(* Logix 5000 project; controller _1407974_PSG_7315 vendor 1 type 14 code 154 rev 20.11; software revision 20.06; part 2 of 4 *)
(* tags used below, declared in another part *)
   AI_L_2_1_FW_Pressure : Analog_Input;
   AI_R_2_0_Pure_Steam_Temperature : Analog_Input;
   Alarm_Emergency_Stop : ALIAS FOR Alarms_Warnings.Latch_Bit[0].0;
   Alarm_Emergency_Stop_Ack : ALIAS FOR Alarms_Warnings.Ack[0].0;
   Alarm_Pure_Steam_High_Temp_Timer : TIMER;
   Alarm_Pure_Steam_High_Temperature : ALIAS FOR Alarms_Warnings.Latch_Bit[0].4;
   Alarm_Pure_Steam_High_Temperature_Ack : ALIAS FOR Alarms_Warnings.Ack[0].4;
   Alarm_Pure_Steam_Temp_Error_Timer : TIMER;
   Alarm_Rupture_Disk_Failure : ALIAS FOR Alarms_Warnings.Latch_Bit[0].1;
   Alarm_Rupture_Disk_Failure_Timer : TIMER;
   Alarm_Rupture_Disk_Faiure_Ack : ALIAS FOR Alarms_Warnings.Ack[0].1;
   Alarm_Separator_High_Level : ALIAS FOR Alarms_Warnings.Latch_Bit[0].2;
   Alarm_Separator_High_Level_Ack : ALIAS FOR Alarms_Warnings.Ack[0].2;
   Alarm_Separator_High_Level_Timer : TIMER;
   Alarm_Separator_Low_Level : ALIAS FOR Alarms_Warnings.Latch_Bit[0].3;
   Alarm_Separator_Low_Level_Ack : ALIAS FOR Alarms_Warnings.Ack[0].3;
   Alarm_Separator_Low_Level_Timer_A : TIMER;
   Alarm_Separator_Low_Level_Timer_B : TIMER;
   Alarms_Warnings : AW;
   AO_L_3_0_VFD_SPEED : Analog_Output;
   AO_R_4_0_Pure_Steam_Temperature : Analog_Output;
   Calculated_CV_Max_Value : REAL;
   Condensed_Pure_Steam_Warrnings_Disabled : Latched_Push_Button;
   Cooling_State_Latch_Timer : TIMER;
   Cooling_Status_Debounce_Timer : TIMER;
   DI_L_1_0_Emergency_Stop_Relay : ALIAS FOR DI_Local_1.0;
   DI_R_1_0_Hi_Hi_Level_LSHH_1950 : ALIAS FOR DI_Remote_1.0;
   DI_R_1_1_Hi_Level_LSH_1950 : ALIAS FOR DI_Remote_1.1;
   DI_R_1_2_Mid_Level_LSM_1950 : ALIAS FOR DI_Remote_1.2;
   DI_R_1_3_Low_Level_LSL_1950 : ALIAS FOR DI_Remote_1.3;
   DI_R_1_5_Burst_Disk_Sensor_PSH_5820 : ALIAS FOR DI_Remote_1.5;
   DO_L_1_0_Alarm_Relay_Coil : Discrete_Out;
   DO_L_1_10_Available : Discrete_Out;
   DO_L_1_11_Available : Discrete_Out;
   DO_L_1_12_Available : Discrete_Out;
   DO_L_1_13_Available : Discrete_Out;
   DO_L_1_14_Feed_Water_Pump_Contactor : Discrete_Out;
   DO_L_1_15_Feed_Water_Pump_On_Light : Discrete_Out;
   DO_L_1_1_Alarm_Horn : Discrete_Out;
   DO_L_1_2_Alarm_Light : Discrete_Out;
   DO_L_1_3_Ready_Light : Discrete_Out;
   DO_L_1_4_Running_Light : Discrete_Out;
   DO_L_1_5_Hour_Meter : Discrete_Out;
   DO_L_1_6_Available : Discrete_Out;
   DO_L_1_7_Available : Discrete_Out;
   DO_L_1_8_Available : Discrete_Out;
   DO_L_1_9_Available : Discrete_Out;
   DO_R_3_0_Pure_Steam_Temp_Control_YV_4110 : Discrete_Out;
   DO_R_3_1_Primary_Level_Control_YV_4760 : Discrete_Out;
   DO_R_3_2_Secondary_Level_Control_YV_4770 : Discrete_Out;
   DO_R_3_3_Coolant_Shutoff_FCV_3025 : Discrete_Out;
   DO_R_3_4_Degasser_Vent_YV_4255 : Discrete_Out;
   DO_R_3_5_FDW_TR : Discrete_Out;
   DO_R_3_6_Available : Discrete_Out;
   DO_R_3_7_Available : Discrete_Out;
   Feedwater_Pressure_PID : PID;
   Feedwater_Pressure_PID_Auto_Mode : Push_Button;
   Feedwater_Pressure_PID_Manual_Mode : Push_Button;
   Lamp_Test : Push_Button;
   Local_Remote : Latched_Push_Button;
   Low_Level_Latch : BOOL;
   Maintenance_Mode : Latched_Push_Button;
   Network_Start : BOOL;
   Network_Stop : BOOL;
   OIT : OIT_Connections;
   PID_Auto_Mode : Push_Button;
   PID_CV_Max_Value_Initialize : BOOL;
   PID_Loop_Trigger_Timer : TIMER;
   PID_Manual_Mode : Push_Button;
   PID_Ramp_Timer : TIMER;
   PS_Temp_GEQ_SetPoint_Minus_5_Deg : BOOL;
   PS_Temp_Setpoint_Minus_5_Deg : REAL;
   Pure_Steam_Temp_Output_Clamp : BOOL;
   Pure_Steam_Temperature : PID;
   Start : Push_Button;
   Stop : Push_Button;
   Unit_Hot : BOOL;
   Unit_Status : Unit_Status;
(* MainProgram, continued *)

ROUTINE _050_Maintenance   (* ladder *)
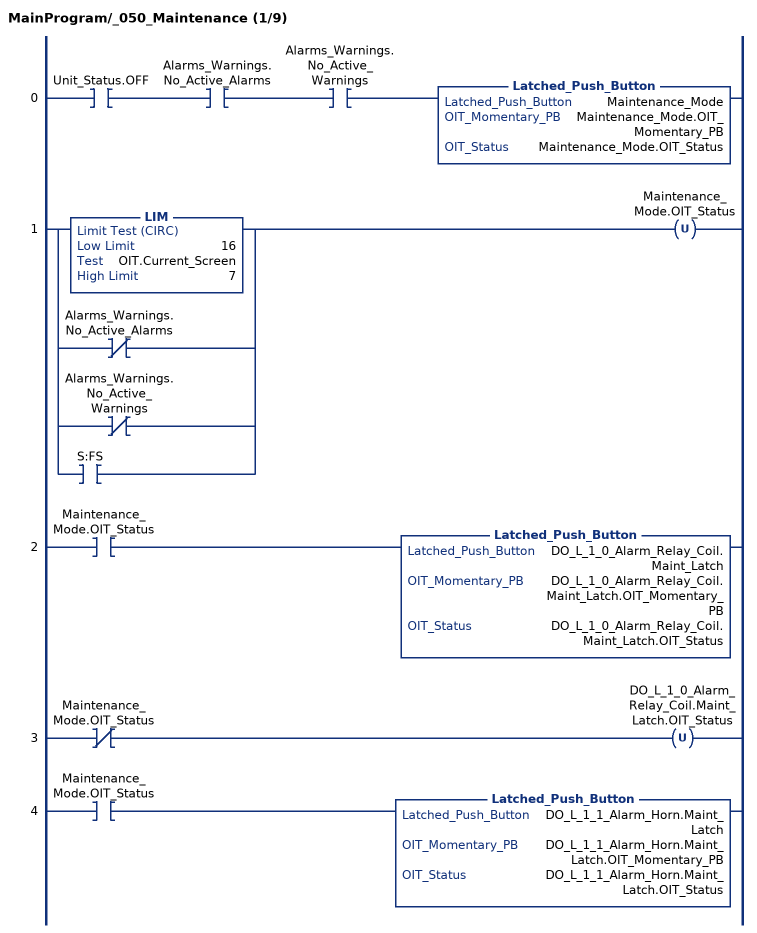
   0: XIC(Unit_Status.OFF)XIC(Alarms_Warnings.No_Active_Alarms)XIC(Alarms_Warnings.No_Active_Warnings)Latched_Push_Button(Maintenance_Mode,Maintenance_Mode.OIT_Momentary_PB,Maintenance_Mode.OIT_Status);
   1: [LIM(16,OIT.Current_Screen,7) ,XIO(Alarms_Warnings.No_Active_Alarms) ,XIO(Alarms_Warnings.No_Active_Warnings) ,XIC(S:FS) ]OTU(Maintenance_Mode.OIT_Status);
   2: XIC(Maintenance_Mode.OIT_Status)Latched_Push_Button(DO_L_1_0_Alarm_Relay_Coil.Maint_Latch,DO_L_1_0_Alarm_Relay_Coil.Maint_Latch.OIT_Momentary_PB,DO_L_1_0_Alarm_Relay_Coil.Maint_Latch.OIT_Status);
   3: XIO(Maintenance_Mode.OIT_Status)OTU(DO_L_1_0_Alarm_Relay_Coil.Maint_Latch.OIT_Status);
   4: XIC(Maintenance_Mode.OIT_Status)Latched_Push_Button(DO_L_1_1_Alarm_Horn.Maint_Latch,DO_L_1_1_Alarm_Horn.Maint_Latch.OIT_Momentary_PB,DO_L_1_1_Alarm_Horn.Maint_Latch.OIT_Status);
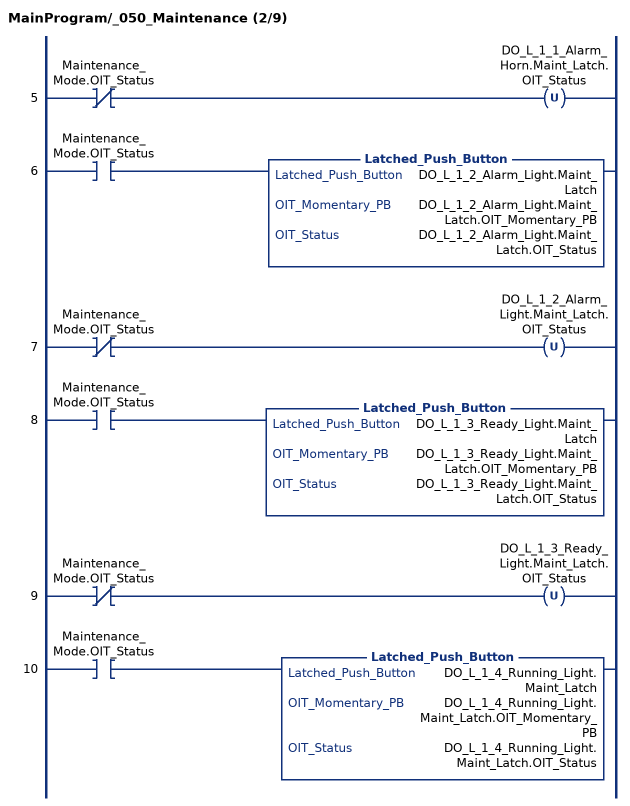
   5: XIO(Maintenance_Mode.OIT_Status)OTU(DO_L_1_1_Alarm_Horn.Maint_Latch.OIT_Status);
   6: XIC(Maintenance_Mode.OIT_Status)Latched_Push_Button(DO_L_1_2_Alarm_Light.Maint_Latch,DO_L_1_2_Alarm_Light.Maint_Latch.OIT_Momentary_PB,DO_L_1_2_Alarm_Light.Maint_Latch.OIT_Status);
   7: XIO(Maintenance_Mode.OIT_Status)OTU(DO_L_1_2_Alarm_Light.Maint_Latch.OIT_Status);
   8: XIC(Maintenance_Mode.OIT_Status)Latched_Push_Button(DO_L_1_3_Ready_Light.Maint_Latch,DO_L_1_3_Ready_Light.Maint_Latch.OIT_Momentary_PB,DO_L_1_3_Ready_Light.Maint_Latch.OIT_Status);
   9: XIO(Maintenance_Mode.OIT_Status)OTU(DO_L_1_3_Ready_Light.Maint_Latch.OIT_Status);
   10: XIC(Maintenance_Mode.OIT_Status)Latched_Push_Button(DO_L_1_4_Running_Light.Maint_Latch,DO_L_1_4_Running_Light.Maint_Latch.OIT_Momentary_PB,DO_L_1_4_Running_Light.Maint_Latch.OIT_Status);
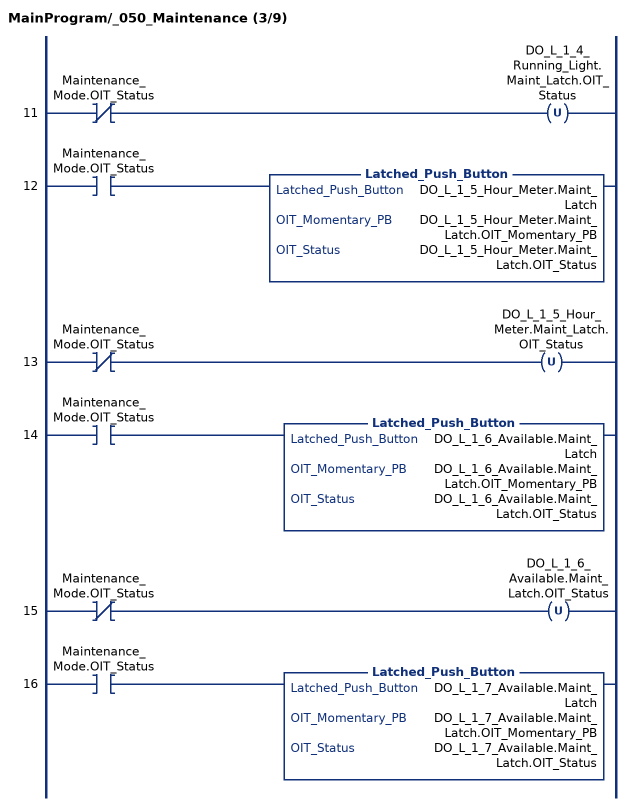
   11: XIO(Maintenance_Mode.OIT_Status)OTU(DO_L_1_4_Running_Light.Maint_Latch.OIT_Status);
   12: XIC(Maintenance_Mode.OIT_Status)Latched_Push_Button(DO_L_1_5_Hour_Meter.Maint_Latch,DO_L_1_5_Hour_Meter.Maint_Latch.OIT_Momentary_PB,DO_L_1_5_Hour_Meter.Maint_Latch.OIT_Status);
   13: XIO(Maintenance_Mode.OIT_Status)OTU(DO_L_1_5_Hour_Meter.Maint_Latch.OIT_Status);
   14: XIC(Maintenance_Mode.OIT_Status)Latched_Push_Button(DO_L_1_6_Available.Maint_Latch,DO_L_1_6_Available.Maint_Latch.OIT_Momentary_PB,DO_L_1_6_Available.Maint_Latch.OIT_Status);
   15: XIO(Maintenance_Mode.OIT_Status)OTU(DO_L_1_6_Available.Maint_Latch.OIT_Status);
   16: XIC(Maintenance_Mode.OIT_Status)Latched_Push_Button(DO_L_1_7_Available.Maint_Latch,DO_L_1_7_Available.Maint_Latch.OIT_Momentary_PB,DO_L_1_7_Available.Maint_Latch.OIT_Status);
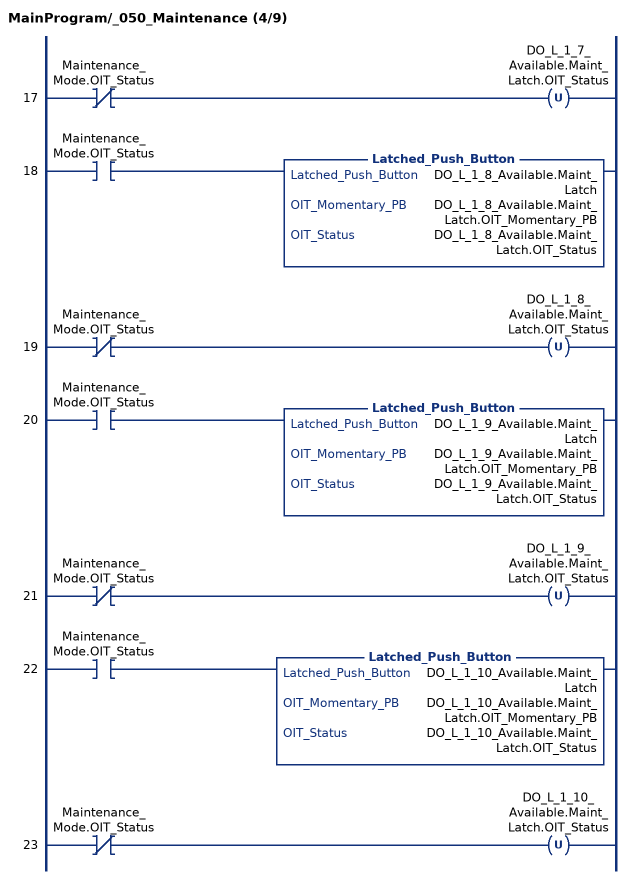
   17: XIO(Maintenance_Mode.OIT_Status)OTU(DO_L_1_7_Available.Maint_Latch.OIT_Status);
   18: XIC(Maintenance_Mode.OIT_Status)Latched_Push_Button(DO_L_1_8_Available.Maint_Latch,DO_L_1_8_Available.Maint_Latch.OIT_Momentary_PB,DO_L_1_8_Available.Maint_Latch.OIT_Status);
   19: XIO(Maintenance_Mode.OIT_Status)OTU(DO_L_1_8_Available.Maint_Latch.OIT_Status);
   20: XIC(Maintenance_Mode.OIT_Status)Latched_Push_Button(DO_L_1_9_Available.Maint_Latch,DO_L_1_9_Available.Maint_Latch.OIT_Momentary_PB,DO_L_1_9_Available.Maint_Latch.OIT_Status);
   21: XIO(Maintenance_Mode.OIT_Status)OTU(DO_L_1_9_Available.Maint_Latch.OIT_Status);
   22: XIC(Maintenance_Mode.OIT_Status)Latched_Push_Button(DO_L_1_10_Available.Maint_Latch,DO_L_1_10_Available.Maint_Latch.OIT_Momentary_PB,DO_L_1_10_Available.Maint_Latch.OIT_Status);
   23: XIO(Maintenance_Mode.OIT_Status)OTU(DO_L_1_10_Available.Maint_Latch.OIT_Status);
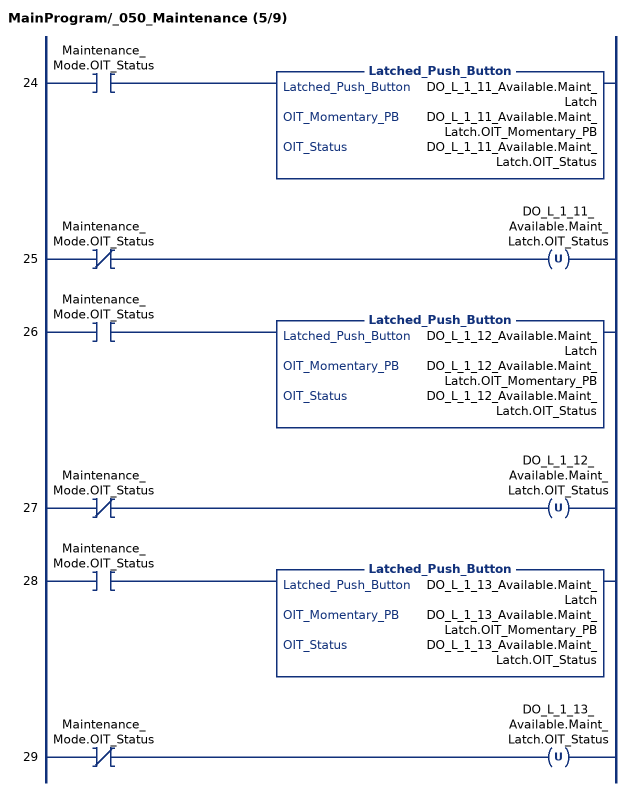
   24: XIC(Maintenance_Mode.OIT_Status)Latched_Push_Button(DO_L_1_11_Available.Maint_Latch,DO_L_1_11_Available.Maint_Latch.OIT_Momentary_PB,DO_L_1_11_Available.Maint_Latch.OIT_Status);
   25: XIO(Maintenance_Mode.OIT_Status)OTU(DO_L_1_11_Available.Maint_Latch.OIT_Status);
   26: XIC(Maintenance_Mode.OIT_Status)Latched_Push_Button(DO_L_1_12_Available.Maint_Latch,DO_L_1_12_Available.Maint_Latch.OIT_Momentary_PB,DO_L_1_12_Available.Maint_Latch.OIT_Status);
   27: XIO(Maintenance_Mode.OIT_Status)OTU(DO_L_1_12_Available.Maint_Latch.OIT_Status);
   28: XIC(Maintenance_Mode.OIT_Status)Latched_Push_Button(DO_L_1_13_Available.Maint_Latch,DO_L_1_13_Available.Maint_Latch.OIT_Momentary_PB,DO_L_1_13_Available.Maint_Latch.OIT_Status);
   29: XIO(Maintenance_Mode.OIT_Status)OTU(DO_L_1_13_Available.Maint_Latch.OIT_Status);
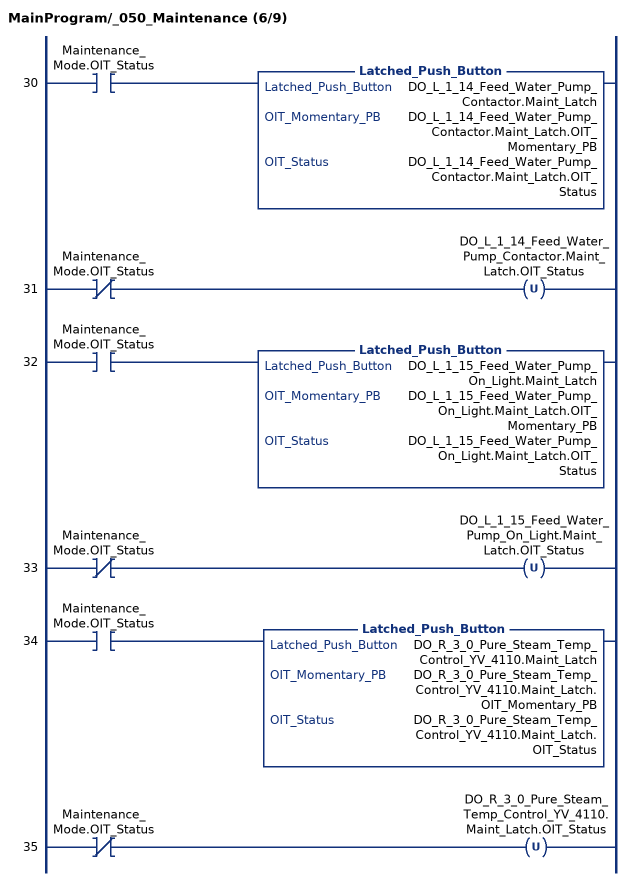
   30: XIC(Maintenance_Mode.OIT_Status)Latched_Push_Button(DO_L_1_14_Feed_Water_Pump_Contactor.Maint_Latch,DO_L_1_14_Feed_Water_Pump_Contactor.Maint_Latch.OIT_Momentary_PB,DO_L_1_14_Feed_Water_Pump_Contactor.Maint_Latch.OIT_Status);
   31: XIO(Maintenance_Mode.OIT_Status)OTU(DO_L_1_14_Feed_Water_Pump_Contactor.Maint_Latch.OIT_Status);
   32: XIC(Maintenance_Mode.OIT_Status)Latched_Push_Button(DO_L_1_15_Feed_Water_Pump_On_Light.Maint_Latch,DO_L_1_15_Feed_Water_Pump_On_Light.Maint_Latch.OIT_Momentary_PB,DO_L_1_15_Feed_Water_Pump_On_Light.Maint_Latch.OIT_Status);
   33: XIO(Maintenance_Mode.OIT_Status)OTU(DO_L_1_15_Feed_Water_Pump_On_Light.Maint_Latch.OIT_Status);
   34: XIC(Maintenance_Mode.OIT_Status)Latched_Push_Button(DO_R_3_0_Pure_Steam_Temp_Control_YV_4110.Maint_Latch,DO_R_3_0_Pure_Steam_Temp_Control_YV_4110.Maint_Latch.OIT_Momentary_PB,DO_R_3_0_Pure_Steam_Temp_Control_YV_4110.Maint_Latch.OIT_Status);
   35: XIO(Maintenance_Mode.OIT_Status)OTU(DO_R_3_0_Pure_Steam_Temp_Control_YV_4110.Maint_Latch.OIT_Status);
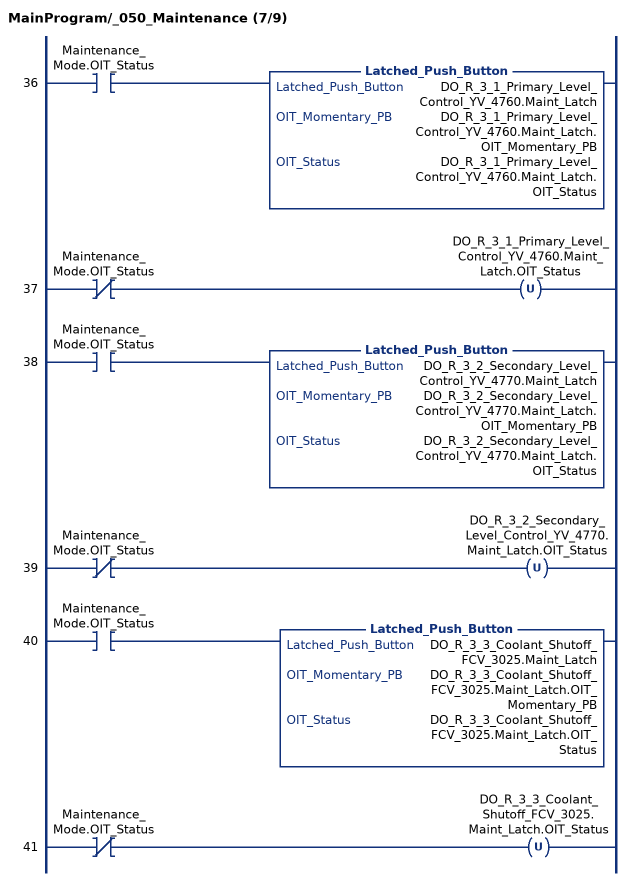
   36: XIC(Maintenance_Mode.OIT_Status)Latched_Push_Button(DO_R_3_1_Primary_Level_Control_YV_4760.Maint_Latch,DO_R_3_1_Primary_Level_Control_YV_4760.Maint_Latch.OIT_Momentary_PB,DO_R_3_1_Primary_Level_Control_YV_4760.Maint_Latch.OIT_Status);
   37: XIO(Maintenance_Mode.OIT_Status)OTU(DO_R_3_1_Primary_Level_Control_YV_4760.Maint_Latch.OIT_Status);
   38: XIC(Maintenance_Mode.OIT_Status)Latched_Push_Button(DO_R_3_2_Secondary_Level_Control_YV_4770.Maint_Latch,DO_R_3_2_Secondary_Level_Control_YV_4770.Maint_Latch.OIT_Momentary_PB,DO_R_3_2_Secondary_Level_Control_YV_4770.Maint_Latch.OIT_Status);
   39: XIO(Maintenance_Mode.OIT_Status)OTU(DO_R_3_2_Secondary_Level_Control_YV_4770.Maint_Latch.OIT_Status);
   40: XIC(Maintenance_Mode.OIT_Status)Latched_Push_Button(DO_R_3_3_Coolant_Shutoff_FCV_3025.Maint_Latch,DO_R_3_3_Coolant_Shutoff_FCV_3025.Maint_Latch.OIT_Momentary_PB,DO_R_3_3_Coolant_Shutoff_FCV_3025.Maint_Latch.OIT_Status);
   41: XIO(Maintenance_Mode.OIT_Status)OTU(DO_R_3_3_Coolant_Shutoff_FCV_3025.Maint_Latch.OIT_Status);
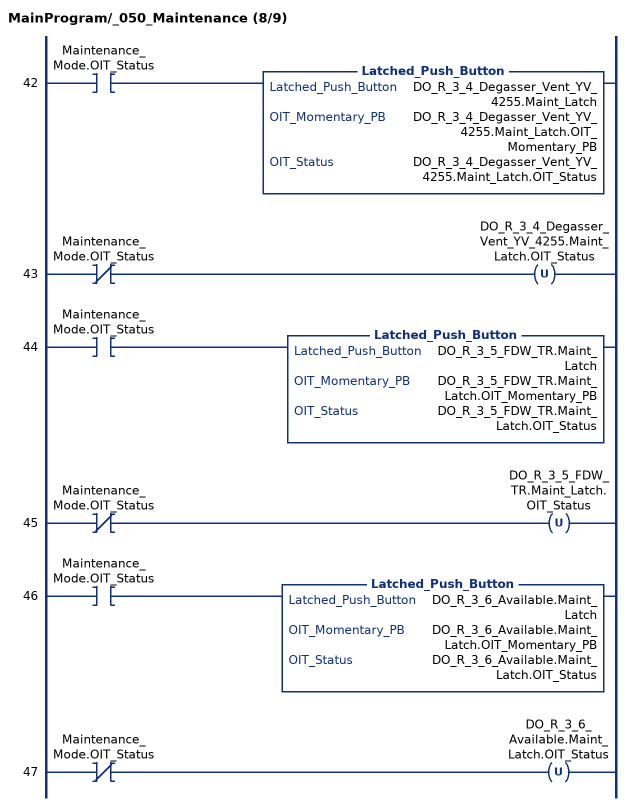
   42: XIC(Maintenance_Mode.OIT_Status)Latched_Push_Button(DO_R_3_4_Degasser_Vent_YV_4255.Maint_Latch,DO_R_3_4_Degasser_Vent_YV_4255.Maint_Latch.OIT_Momentary_PB,DO_R_3_4_Degasser_Vent_YV_4255.Maint_Latch.OIT_Status);
   43: XIO(Maintenance_Mode.OIT_Status)OTU(DO_R_3_4_Degasser_Vent_YV_4255.Maint_Latch.OIT_Status);
   44: XIC(Maintenance_Mode.OIT_Status)Latched_Push_Button(DO_R_3_5_FDW_TR.Maint_Latch,DO_R_3_5_FDW_TR.Maint_Latch.OIT_Momentary_PB,DO_R_3_5_FDW_TR.Maint_Latch.OIT_Status);
   45: XIO(Maintenance_Mode.OIT_Status)OTU(DO_R_3_5_FDW_TR.Maint_Latch.OIT_Status);
   46: XIC(Maintenance_Mode.OIT_Status)Latched_Push_Button(DO_R_3_6_Available.Maint_Latch,DO_R_3_6_Available.Maint_Latch.OIT_Momentary_PB,DO_R_3_6_Available.Maint_Latch.OIT_Status);
   47: XIO(Maintenance_Mode.OIT_Status)OTU(DO_R_3_6_Available.Maint_Latch.OIT_Status);
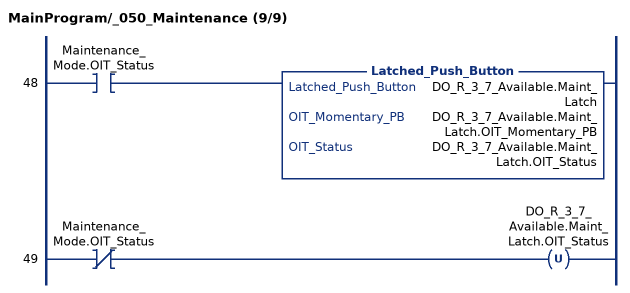
   48: XIC(Maintenance_Mode.OIT_Status)Latched_Push_Button(DO_R_3_7_Available.Maint_Latch,DO_R_3_7_Available.Maint_Latch.OIT_Momentary_PB,DO_R_3_7_Available.Maint_Latch.OIT_Status);
   49: XIO(Maintenance_Mode.OIT_Status)OTU(DO_R_3_7_Available.Maint_Latch.OIT_Status);
END_ROUTINE

ROUTINE _060_Main_Routine   (* ladder *)
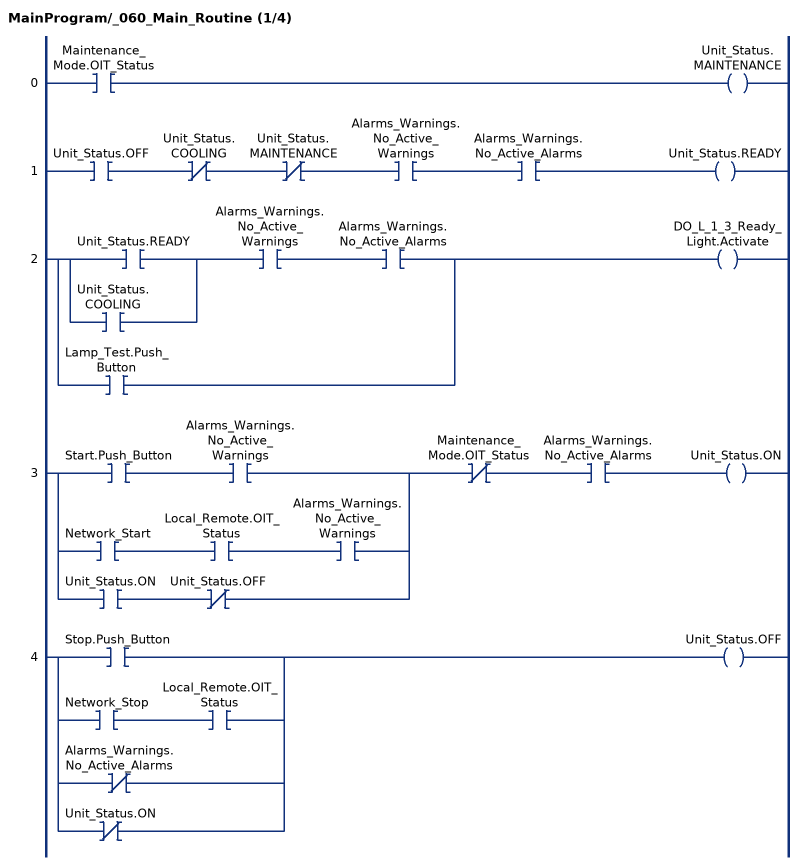
   0: XIC(Maintenance_Mode.OIT_Status)OTE(Unit_Status.MAINTENANCE);
   1: XIC(Unit_Status.OFF)XIO(Unit_Status.COOLING)XIO(Unit_Status.MAINTENANCE)XIC(Alarms_Warnings.No_Active_Warnings)XIC(Alarms_Warnings.No_Active_Alarms)OTE(Unit_Status.READY);
   2: [[XIC(Unit_Status.READY) ,XIC(Unit_Status.COOLING) ] XIC(Alarms_Warnings.No_Active_Warnings) XIC(Alarms_Warnings.No_Active_Alarms) ,XIC(Lamp_Test.Push_Button) ]OTE(DO_L_1_3_Ready_Light.Activate);
   3: [XIC(Start.Push_Button) XIC(Alarms_Warnings.No_Active_Warnings) ,XIC(Network_Start) XIC(Local_Remote.OIT_Status) XIC(Alarms_Warnings.No_Active_Warnings) ,XIC(Unit_Status.ON) XIO(Unit_Status.OFF) ]XIO(Maintenance_Mode.OIT_Status)XIC(Alarms_Warnings.No_Active_Alarms)OTE(Unit_Status.ON);
   4: [XIC(Stop.Push_Button) ,XIC(Network_Stop) XIC(Local_Remote.OIT_Status) ,XIO(Alarms_Warnings.No_Active_Alarms) ,XIO(Unit_Status.ON) ]OTE(Unit_Status.OFF);
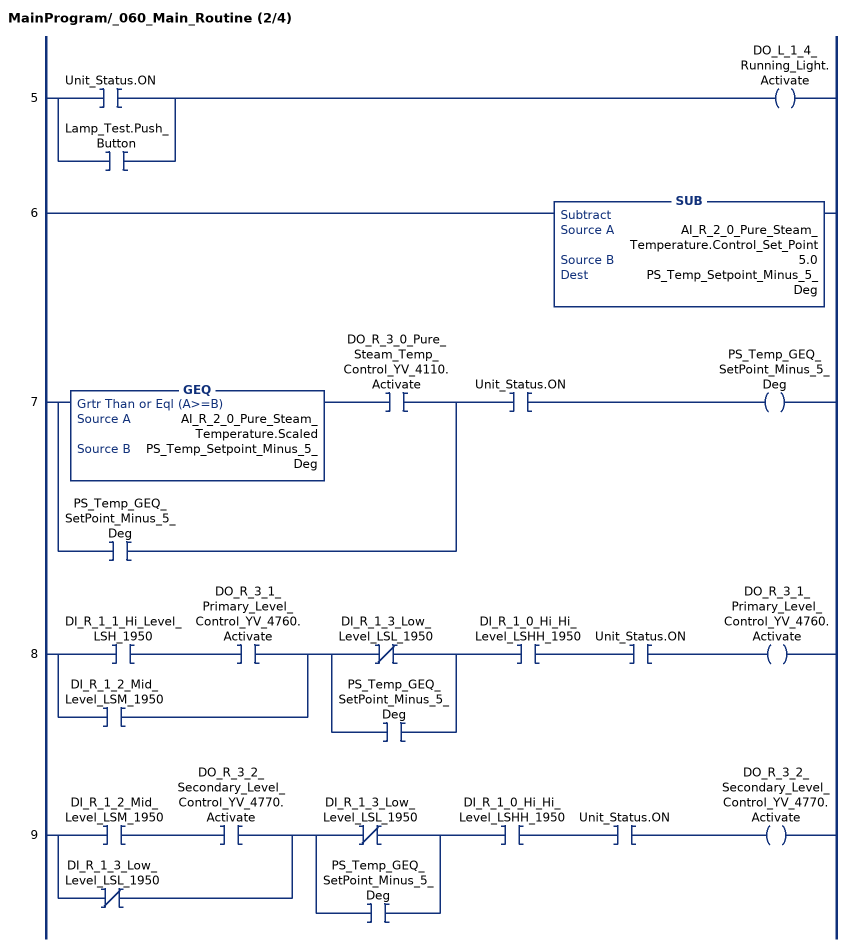
   5: [XIC(Unit_Status.ON) ,XIC(Lamp_Test.Push_Button) ]OTE(DO_L_1_4_Running_Light.Activate);
   6: SUB(AI_R_2_0_Pure_Steam_Temperature.Control_Set_Point,5.0,PS_Temp_Setpoint_Minus_5_Deg);
   7: [GEQ(AI_R_2_0_Pure_Steam_Temperature.Scaled,PS_Temp_Setpoint_Minus_5_Deg) XIC(DO_R_3_0_Pure_Steam_Temp_Control_YV_4110.Activate) ,XIC(PS_Temp_GEQ_SetPoint_Minus_5_Deg) ]XIC(Unit_Status.ON)OTE(PS_Temp_GEQ_SetPoint_Minus_5_Deg);
   8: [XIC(DI_R_1_1_Hi_Level_LSH_1950) XIC(DO_R_3_1_Primary_Level_Control_YV_4760.Activate) ,XIC(DI_R_1_2_Mid_Level_LSM_1950) ][XIO(DI_R_1_3_Low_Level_LSL_1950) ,XIC(PS_Temp_GEQ_SetPoint_Minus_5_Deg) ]XIC(DI_R_1_0_Hi_Hi_Level_LSHH_1950)XIC(Unit_Status.ON)OTE(DO_R_3_1_Primary_Level_Control_YV_4760.Activate);
   9: [XIC(DI_R_1_2_Mid_Level_LSM_1950) XIC(DO_R_3_2_Secondary_Level_Control_YV_4770.Activate) ,XIO(DI_R_1_3_Low_Level_LSL_1950) ][XIO(DI_R_1_3_Low_Level_LSL_1950) ,XIC(PS_Temp_GEQ_SetPoint_Minus_5_Deg) ]XIC(DI_R_1_0_Hi_Hi_Level_LSHH_1950)XIC(Unit_Status.ON)OTE(DO_R_3_2_Secondary_Level_Control_YV_4770.Activate);
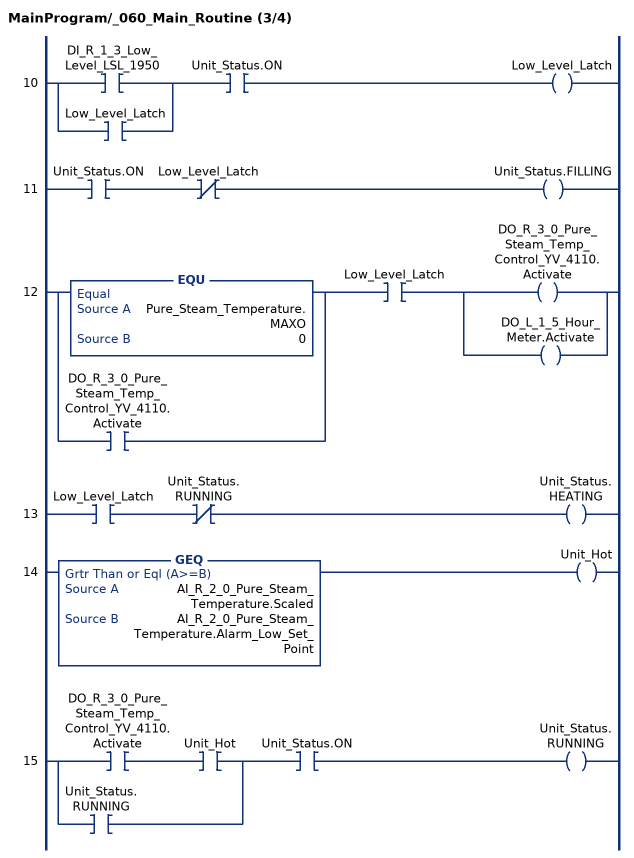
   10: [XIC(DI_R_1_3_Low_Level_LSL_1950) ,XIC(Low_Level_Latch) ]XIC(Unit_Status.ON)OTE(Low_Level_Latch);
   11: XIC(Unit_Status.ON)XIO(Low_Level_Latch)OTE(Unit_Status.FILLING);
   12: [EQU(Pure_Steam_Temperature.MAXO,0) ,XIC(DO_R_3_0_Pure_Steam_Temp_Control_YV_4110.Activate) ]XIC(Low_Level_Latch)[OTE(DO_R_3_0_Pure_Steam_Temp_Control_YV_4110.Activate) ,OTE(DO_L_1_5_Hour_Meter.Activate) ];
   13: XIC(Low_Level_Latch)XIO(Unit_Status.RUNNING)OTE(Unit_Status.HEATING);
   14: GEQ(AI_R_2_0_Pure_Steam_Temperature.Scaled,AI_R_2_0_Pure_Steam_Temperature.Alarm_Low_Set_Point)OTE(Unit_Hot);
   15: [XIC(DO_R_3_0_Pure_Steam_Temp_Control_YV_4110.Activate) XIC(Unit_Hot) ,XIC(Unit_Status.RUNNING) ]XIC(Unit_Status.ON)OTE(Unit_Status.RUNNING);
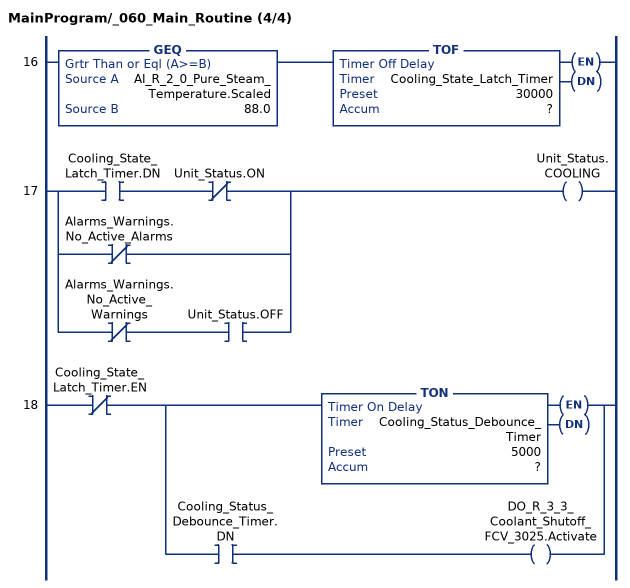
   16: GEQ(AI_R_2_0_Pure_Steam_Temperature.Scaled,88.0)TOF(Cooling_State_Latch_Timer,?,?);
   17: [XIC(Cooling_State_Latch_Timer.DN) XIO(Unit_Status.ON) ,XIO(Alarms_Warnings.No_Active_Alarms) ,XIO(Alarms_Warnings.No_Active_Warnings) XIC(Unit_Status.OFF) ]OTE(Unit_Status.COOLING);
   18: XIO(Cooling_State_Latch_Timer.EN)[TON(Cooling_Status_Debounce_Timer,?,?) ,XIC(Cooling_Status_Debounce_Timer.DN) OTE(DO_R_3_3_Coolant_Shutoff_FCV_3025.Activate) ];
END_ROUTINE

ROUTINE _070_PID   (* ladder *)
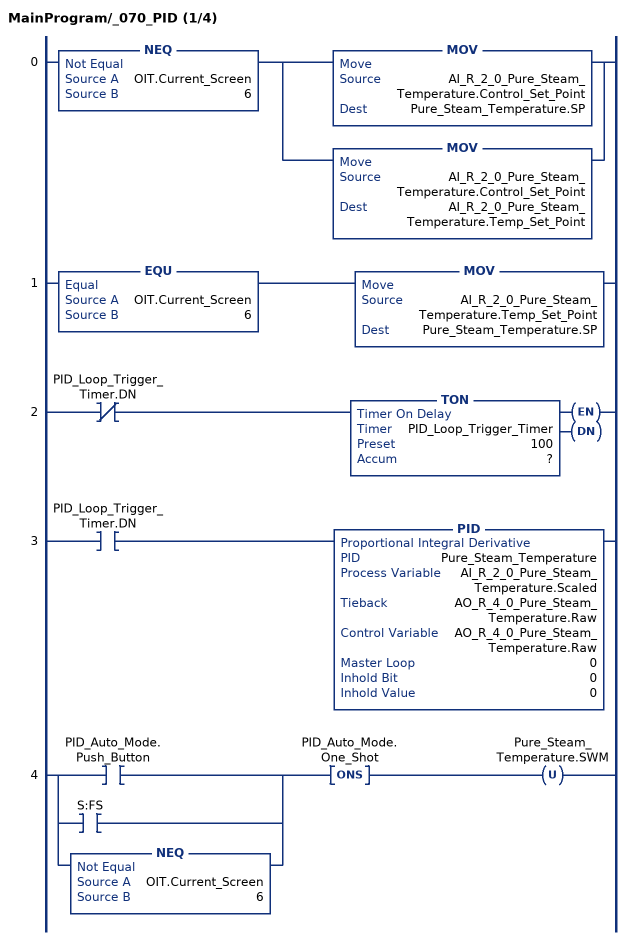
   0: NEQ(OIT.Current_Screen,6)[MOV(AI_R_2_0_Pure_Steam_Temperature.Control_Set_Point,Pure_Steam_Temperature.SP) ,MOV(AI_R_2_0_Pure_Steam_Temperature.Control_Set_Point,AI_R_2_0_Pure_Steam_Temperature.Temp_Set_Point) ];
   1: EQU(OIT.Current_Screen,6)MOV(AI_R_2_0_Pure_Steam_Temperature.Temp_Set_Point,Pure_Steam_Temperature.SP);
   2: XIO(PID_Loop_Trigger_Timer.DN)TON(PID_Loop_Trigger_Timer,?,?);
   3: XIC(PID_Loop_Trigger_Timer.DN)PID(Pure_Steam_Temperature,AI_R_2_0_Pure_Steam_Temperature.Scaled,AO_R_4_0_Pure_Steam_Temperature.Raw,AO_R_4_0_Pure_Steam_Temperature.Raw,0,0,0);
   4: [XIC(PID_Auto_Mode.Push_Button) ,XIC(S:FS) ,NEQ(OIT.Current_Screen,6) ]ONS(PID_Auto_Mode.One_Shot)OTU(Pure_Steam_Temperature.SWM);
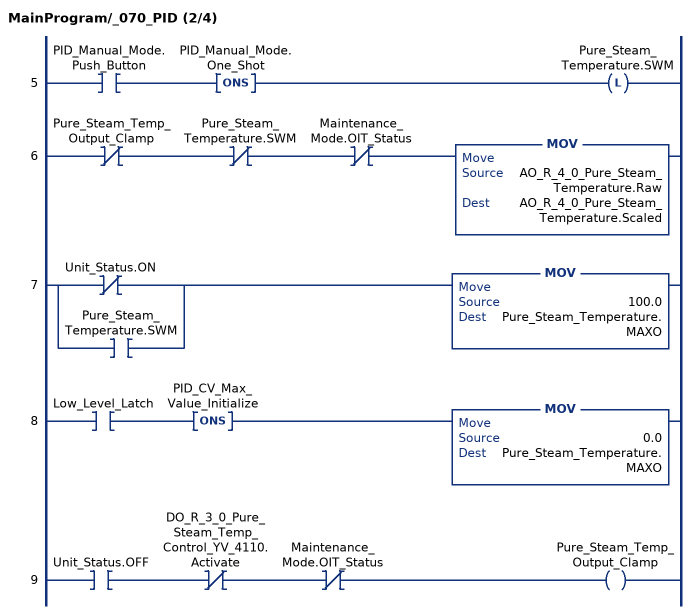
   5: XIC(PID_Manual_Mode.Push_Button)ONS(PID_Manual_Mode.One_Shot)OTL(Pure_Steam_Temperature.SWM);
   6: XIO(Pure_Steam_Temp_Output_Clamp)XIO(Pure_Steam_Temperature.SWM)XIO(Maintenance_Mode.OIT_Status)MOV(AO_R_4_0_Pure_Steam_Temperature.Raw,AO_R_4_0_Pure_Steam_Temperature.Scaled);
   7: [XIO(Unit_Status.ON) ,XIC(Pure_Steam_Temperature.SWM) ]MOV(100.0,Pure_Steam_Temperature.MAXO);
   8: XIC(Low_Level_Latch)ONS(PID_CV_Max_Value_Initialize)MOV(0.0,Pure_Steam_Temperature.MAXO);
   9: XIC(Unit_Status.OFF)XIO(DO_R_3_0_Pure_Steam_Temp_Control_YV_4110.Activate)XIO(Maintenance_Mode.OIT_Status)OTE(Pure_Steam_Temp_Output_Clamp);
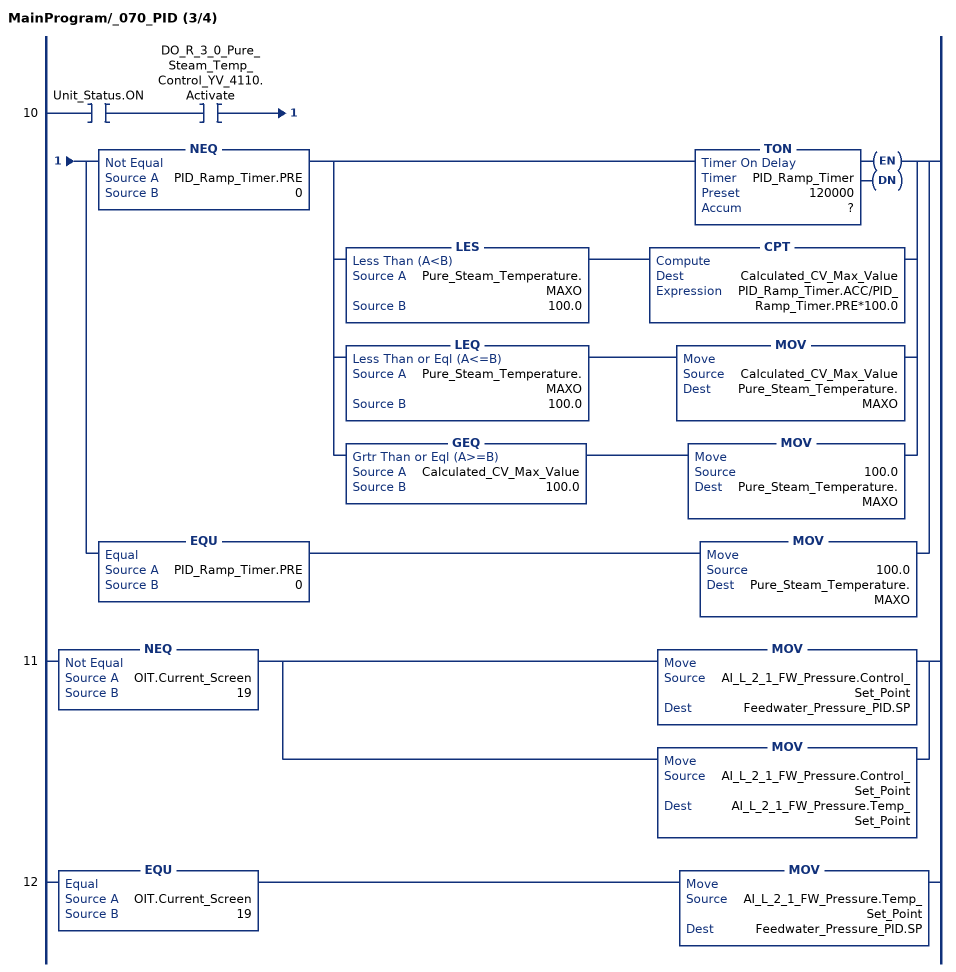
   10: XIC(Unit_Status.ON)XIC(DO_R_3_0_Pure_Steam_Temp_Control_YV_4110.Activate)[NEQ(PID_Ramp_Timer.PRE,0) [TON(PID_Ramp_Timer,?,?) ,LES(Pure_Steam_Temperature.MAXO,100.0) CPT(Calculated_CV_Max_Value,PID_Ramp_Timer.ACC/PID_Ramp_Timer.PRE*100.0) ,LEQ(Pure_Steam_Temperature.MAXO,100.0) MOV(Calculated_CV_Max_Value,Pure_Steam_Temperature.MAXO) ,GEQ(Calculated_CV_Max_Value,100.0) MOV(100.0,Pure_Steam_Temperature.MAXO) ] ,EQU(PID_Ramp_Timer.PRE,0) MOV(100.0,Pure_Steam_Temperature.MAXO) ];
   11: NEQ(OIT.Current_Screen,19)[MOV(AI_L_2_1_FW_Pressure.Control_Set_Point,Feedwater_Pressure_PID.SP) ,MOV(AI_L_2_1_FW_Pressure.Control_Set_Point,AI_L_2_1_FW_Pressure.Temp_Set_Point) ];
   12: EQU(OIT.Current_Screen,19)MOV(AI_L_2_1_FW_Pressure.Temp_Set_Point,Feedwater_Pressure_PID.SP);
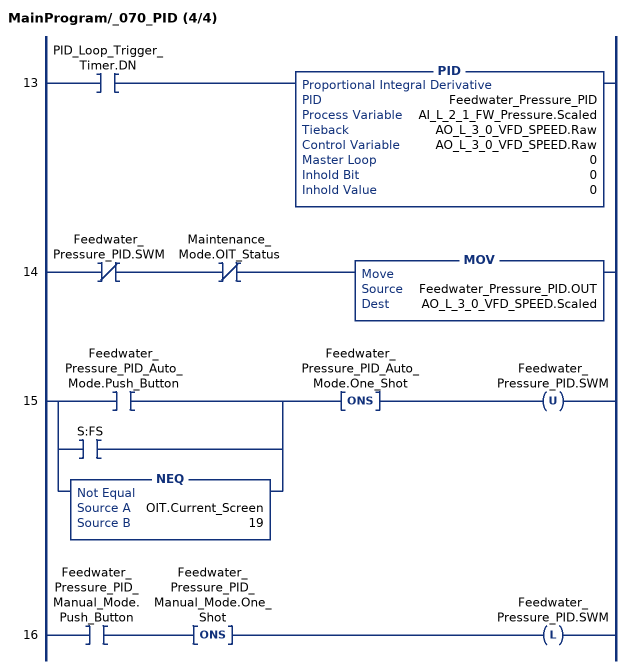
   13: XIC(PID_Loop_Trigger_Timer.DN)PID(Feedwater_Pressure_PID,AI_L_2_1_FW_Pressure.Scaled,AO_L_3_0_VFD_SPEED.Raw,AO_L_3_0_VFD_SPEED.Raw,0,0,0);
   14: XIO(Feedwater_Pressure_PID.SWM)XIO(Maintenance_Mode.OIT_Status)MOV(Feedwater_Pressure_PID.OUT,AO_L_3_0_VFD_SPEED.Scaled);
   15: [XIC(Feedwater_Pressure_PID_Auto_Mode.Push_Button) ,XIC(S:FS) ,NEQ(OIT.Current_Screen,19) ]ONS(Feedwater_Pressure_PID_Auto_Mode.One_Shot)OTU(Feedwater_Pressure_PID.SWM);
   16: XIC(Feedwater_Pressure_PID_Manual_Mode.Push_Button)ONS(Feedwater_Pressure_PID_Manual_Mode.One_Shot)OTL(Feedwater_Pressure_PID.SWM);
END_ROUTINE

ROUTINE _080_Alarms_Warnings   (* ladder *)
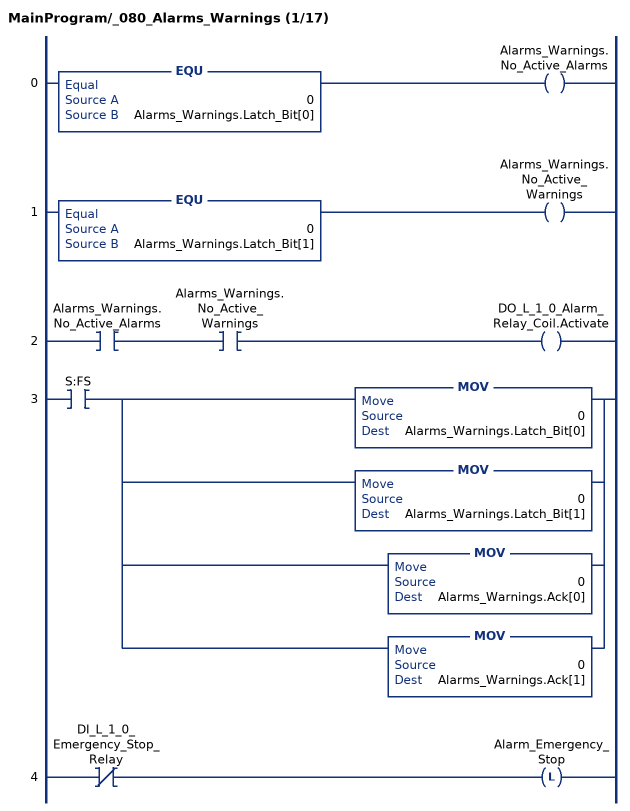
   0: EQU(0,Alarms_Warnings.Latch_Bit[0])OTE(Alarms_Warnings.No_Active_Alarms);
   1: EQU(0,Alarms_Warnings.Latch_Bit[1])OTE(Alarms_Warnings.No_Active_Warnings);
   2: XIC(Alarms_Warnings.No_Active_Alarms)XIC(Alarms_Warnings.No_Active_Warnings)OTE(DO_L_1_0_Alarm_Relay_Coil.Activate);
   3: XIC(S:FS)[MOV(0,Alarms_Warnings.Latch_Bit[0]) ,MOV(0,Alarms_Warnings.Latch_Bit[1]) ,MOV(0,Alarms_Warnings.Ack[0]) ,MOV(0,Alarms_Warnings.Ack[1]) ];
   4: XIO(DI_L_1_0_Emergency_Stop_Relay)OTL(Alarm_Emergency_Stop);
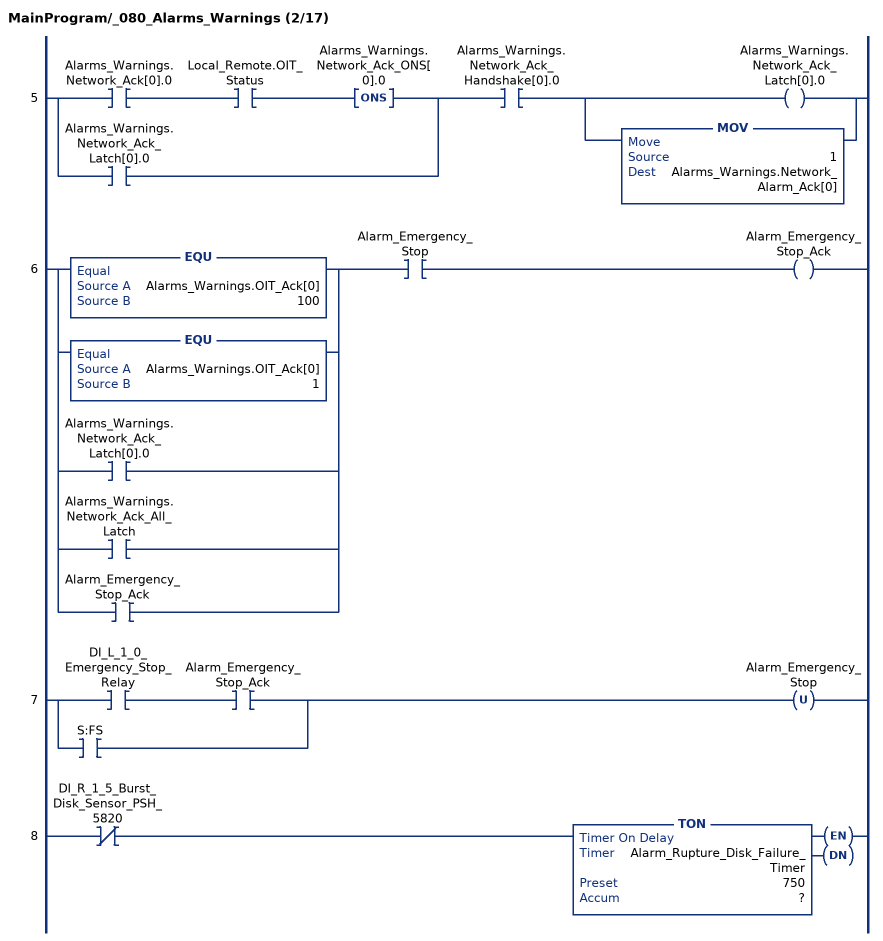
   5: [XIC(Alarms_Warnings.Network_Ack[0].0) XIC(Local_Remote.OIT_Status) ONS(Alarms_Warnings.Network_Ack_ONS[0].0) ,XIC(Alarms_Warnings.Network_Ack_Latch[0].0) ]XIC(Alarms_Warnings.Network_Ack_Handshake[0].0)[OTE(Alarms_Warnings.Network_Ack_Latch[0].0) ,MOV(1,Alarms_Warnings.Network_Alarm_Ack[0]) ];
   6: [EQU(Alarms_Warnings.OIT_Ack[0],100) ,EQU(Alarms_Warnings.OIT_Ack[0],1) ,XIC(Alarms_Warnings.Network_Ack_Latch[0].0) ,XIC(Alarms_Warnings.Network_Ack_All_Latch) ,XIC(Alarm_Emergency_Stop_Ack) ]XIC(Alarm_Emergency_Stop)OTE(Alarm_Emergency_Stop_Ack);
   7: [XIC(DI_L_1_0_Emergency_Stop_Relay) XIC(Alarm_Emergency_Stop_Ack) ,XIC(S:FS) ]OTU(Alarm_Emergency_Stop);
   8: XIO(DI_R_1_5_Burst_Disk_Sensor_PSH_5820)TON(Alarm_Rupture_Disk_Failure_Timer,?,?);
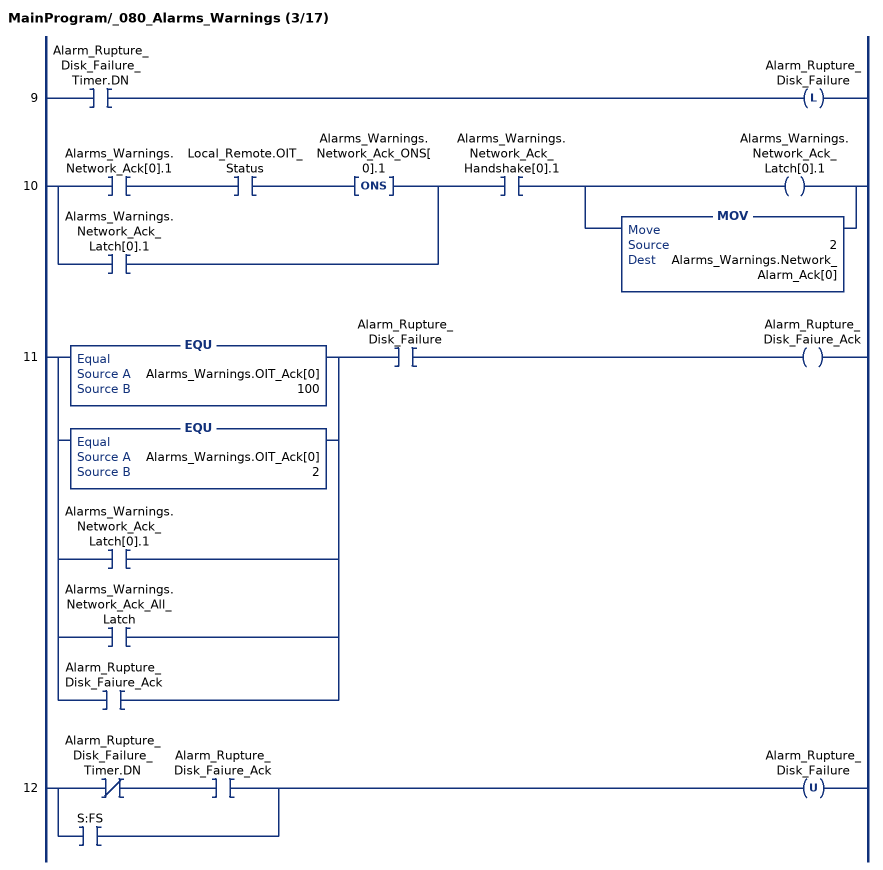
   9: XIC(Alarm_Rupture_Disk_Failure_Timer.DN)OTL(Alarm_Rupture_Disk_Failure);
   10: [XIC(Alarms_Warnings.Network_Ack[0].1) XIC(Local_Remote.OIT_Status) ONS(Alarms_Warnings.Network_Ack_ONS[0].1) ,XIC(Alarms_Warnings.Network_Ack_Latch[0].1) ]XIC(Alarms_Warnings.Network_Ack_Handshake[0].1)[OTE(Alarms_Warnings.Network_Ack_Latch[0].1) ,MOV(2,Alarms_Warnings.Network_Alarm_Ack[0]) ];
   11: [EQU(Alarms_Warnings.OIT_Ack[0],100) ,EQU(Alarms_Warnings.OIT_Ack[0],2) ,XIC(Alarms_Warnings.Network_Ack_Latch[0].1) ,XIC(Alarms_Warnings.Network_Ack_All_Latch) ,XIC(Alarm_Rupture_Disk_Faiure_Ack) ]XIC(Alarm_Rupture_Disk_Failure)OTE(Alarm_Rupture_Disk_Faiure_Ack);
   12: [XIO(Alarm_Rupture_Disk_Failure_Timer.DN) XIC(Alarm_Rupture_Disk_Faiure_Ack) ,XIC(S:FS) ]OTU(Alarm_Rupture_Disk_Failure);
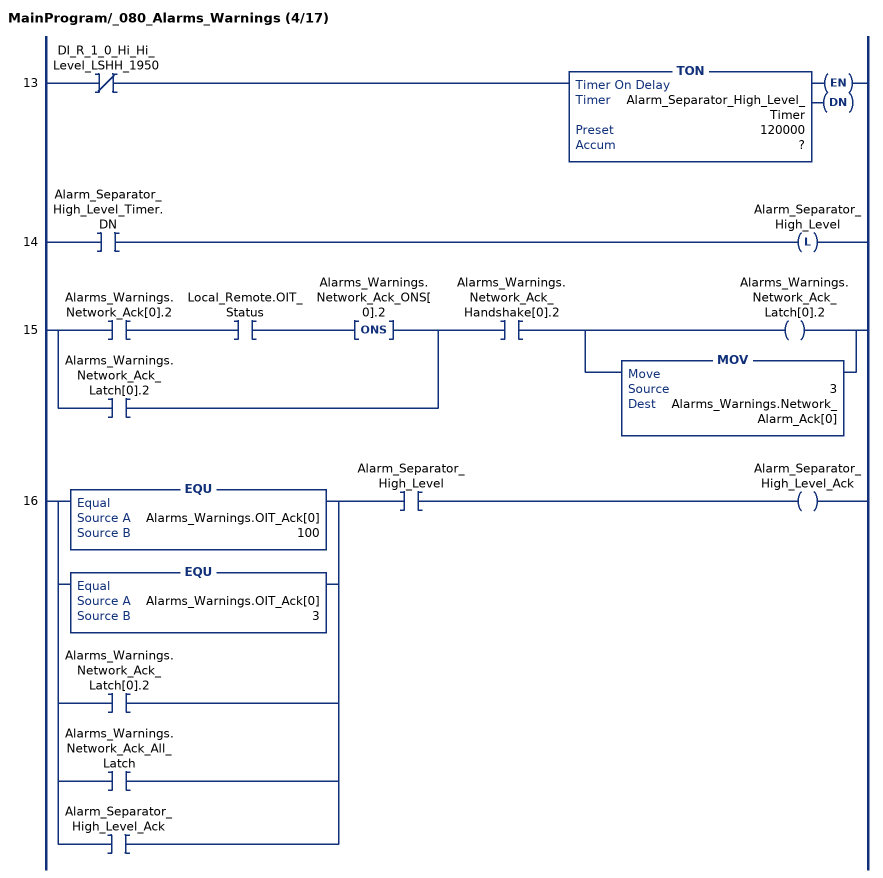
   13: XIO(DI_R_1_0_Hi_Hi_Level_LSHH_1950)TON(Alarm_Separator_High_Level_Timer,?,?);
   14: XIC(Alarm_Separator_High_Level_Timer.DN)OTL(Alarm_Separator_High_Level);
   15: [XIC(Alarms_Warnings.Network_Ack[0].2) XIC(Local_Remote.OIT_Status) ONS(Alarms_Warnings.Network_Ack_ONS[0].2) ,XIC(Alarms_Warnings.Network_Ack_Latch[0].2) ]XIC(Alarms_Warnings.Network_Ack_Handshake[0].2)[OTE(Alarms_Warnings.Network_Ack_Latch[0].2) ,MOV(3,Alarms_Warnings.Network_Alarm_Ack[0]) ];
   16: [EQU(Alarms_Warnings.OIT_Ack[0],100) ,EQU(Alarms_Warnings.OIT_Ack[0],3) ,XIC(Alarms_Warnings.Network_Ack_Latch[0].2) ,XIC(Alarms_Warnings.Network_Ack_All_Latch) ,XIC(Alarm_Separator_High_Level_Ack) ]XIC(Alarm_Separator_High_Level)OTE(Alarm_Separator_High_Level_Ack);
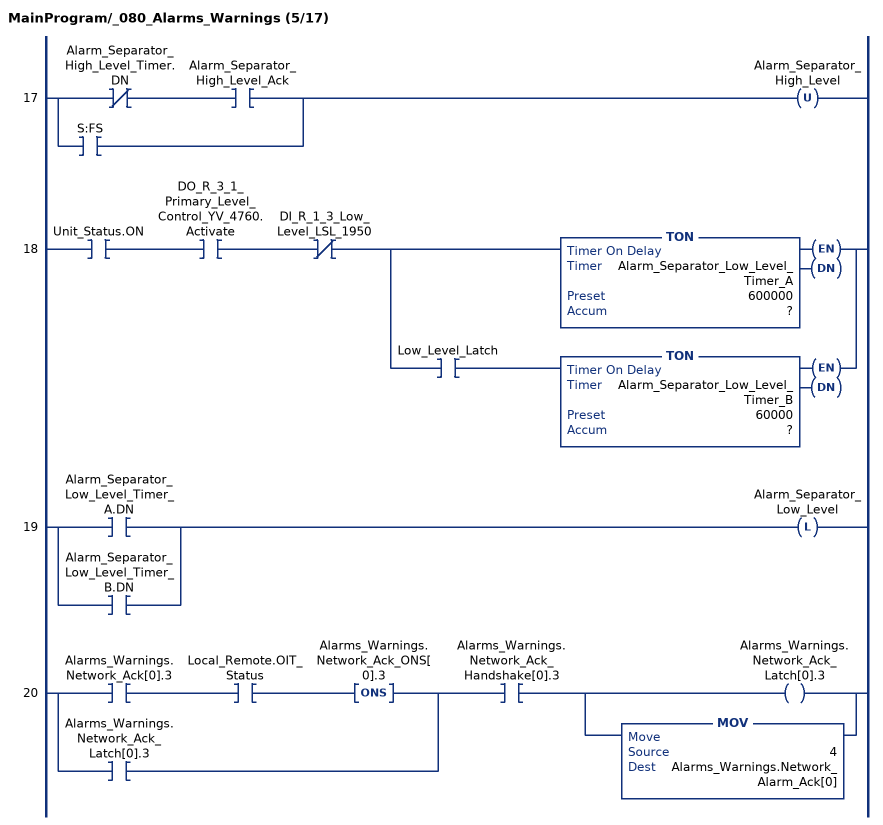
   17: [XIO(Alarm_Separator_High_Level_Timer.DN) XIC(Alarm_Separator_High_Level_Ack) ,XIC(S:FS) ]OTU(Alarm_Separator_High_Level);
   18: XIC(Unit_Status.ON)XIC(DO_R_3_1_Primary_Level_Control_YV_4760.Activate)XIO(DI_R_1_3_Low_Level_LSL_1950)[TON(Alarm_Separator_Low_Level_Timer_A,?,?) ,XIC(Low_Level_Latch) TON(Alarm_Separator_Low_Level_Timer_B,?,?) ];
   19: [XIC(Alarm_Separator_Low_Level_Timer_A.DN) ,XIC(Alarm_Separator_Low_Level_Timer_B.DN) ]OTL(Alarm_Separator_Low_Level);
   20: [XIC(Alarms_Warnings.Network_Ack[0].3) XIC(Local_Remote.OIT_Status) ONS(Alarms_Warnings.Network_Ack_ONS[0].3) ,XIC(Alarms_Warnings.Network_Ack_Latch[0].3) ]XIC(Alarms_Warnings.Network_Ack_Handshake[0].3)[OTE(Alarms_Warnings.Network_Ack_Latch[0].3) ,MOV(4,Alarms_Warnings.Network_Alarm_Ack[0]) ];
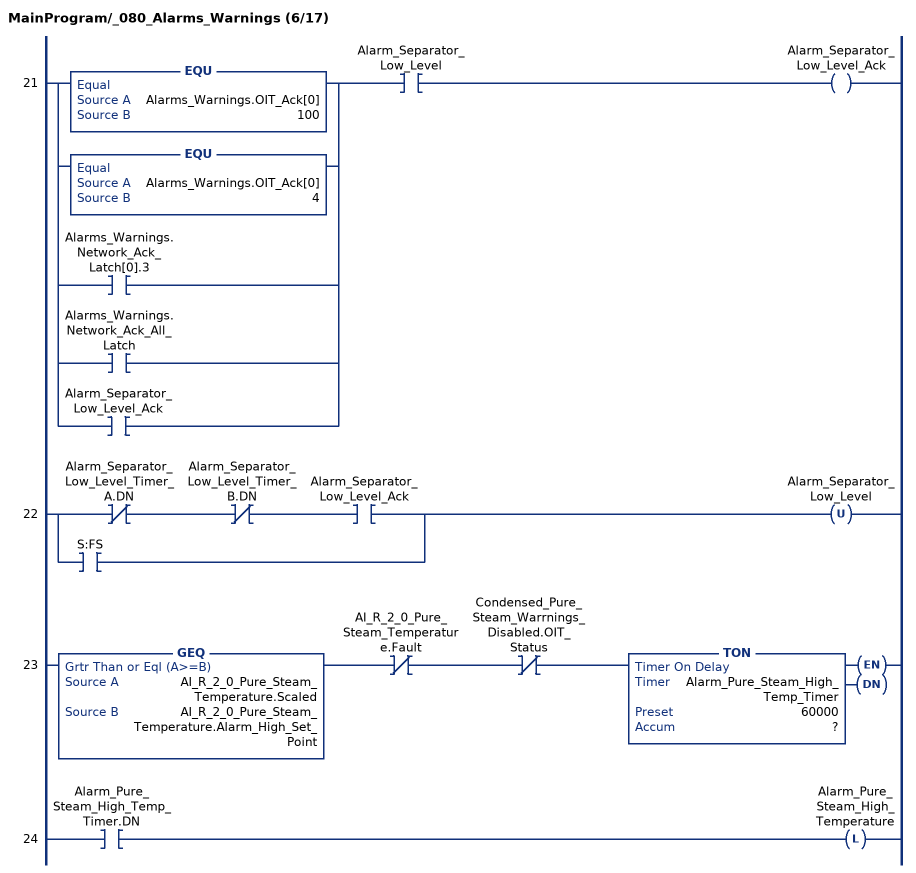
   21: [EQU(Alarms_Warnings.OIT_Ack[0],100) ,EQU(Alarms_Warnings.OIT_Ack[0],4) ,XIC(Alarms_Warnings.Network_Ack_Latch[0].3) ,XIC(Alarms_Warnings.Network_Ack_All_Latch) ,XIC(Alarm_Separator_Low_Level_Ack) ]XIC(Alarm_Separator_Low_Level)OTE(Alarm_Separator_Low_Level_Ack);
   22: [XIO(Alarm_Separator_Low_Level_Timer_A.DN) XIO(Alarm_Separator_Low_Level_Timer_B.DN) XIC(Alarm_Separator_Low_Level_Ack) ,XIC(S:FS) ]OTU(Alarm_Separator_Low_Level);
   23: GEQ(AI_R_2_0_Pure_Steam_Temperature.Scaled,AI_R_2_0_Pure_Steam_Temperature.Alarm_High_Set_Point)XIO(AI_R_2_0_Pure_Steam_Temperature.Fault)XIO(Condensed_Pure_Steam_Warrnings_Disabled.OIT_Status)TON(Alarm_Pure_Steam_High_Temp_Timer,?,?);
   24: XIC(Alarm_Pure_Steam_High_Temp_Timer.DN)OTL(Alarm_Pure_Steam_High_Temperature);
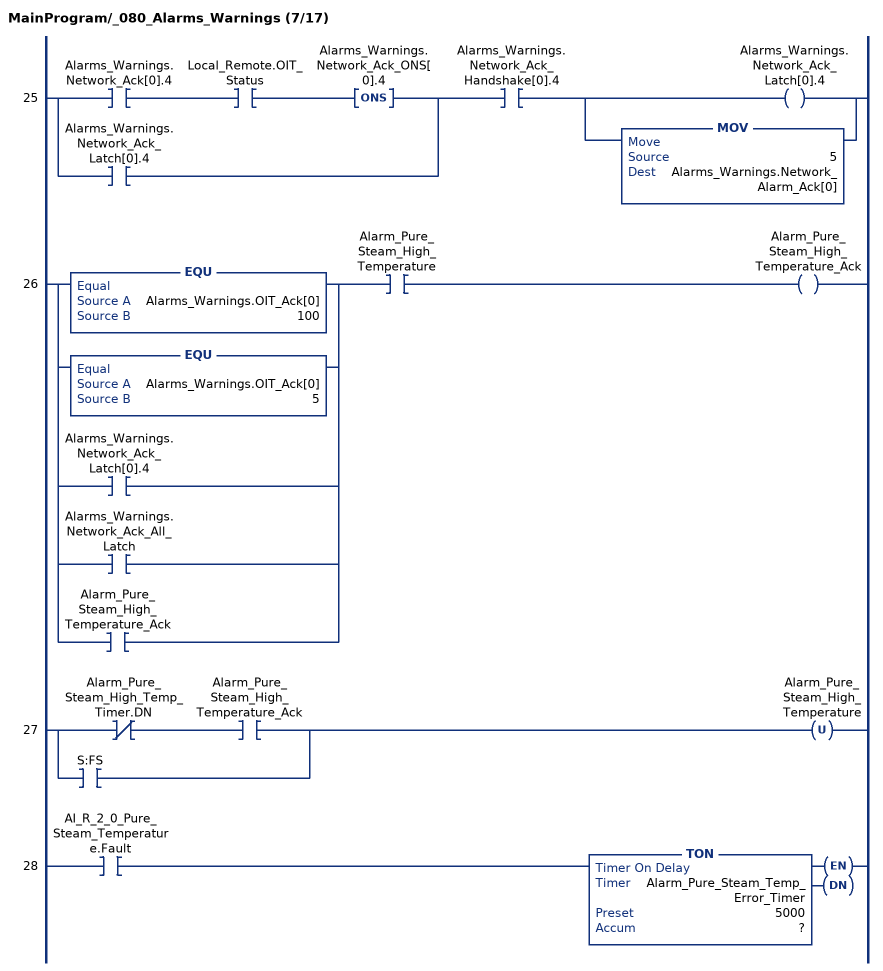
   25: [XIC(Alarms_Warnings.Network_Ack[0].4) XIC(Local_Remote.OIT_Status) ONS(Alarms_Warnings.Network_Ack_ONS[0].4) ,XIC(Alarms_Warnings.Network_Ack_Latch[0].4) ]XIC(Alarms_Warnings.Network_Ack_Handshake[0].4)[OTE(Alarms_Warnings.Network_Ack_Latch[0].4) ,MOV(5,Alarms_Warnings.Network_Alarm_Ack[0]) ];
   26: [EQU(Alarms_Warnings.OIT_Ack[0],100) ,EQU(Alarms_Warnings.OIT_Ack[0],5) ,XIC(Alarms_Warnings.Network_Ack_Latch[0].4) ,XIC(Alarms_Warnings.Network_Ack_All_Latch) ,XIC(Alarm_Pure_Steam_High_Temperature_Ack) ]XIC(Alarm_Pure_Steam_High_Temperature)OTE(Alarm_Pure_Steam_High_Temperature_Ack);
   27: [XIO(Alarm_Pure_Steam_High_Temp_Timer.DN) XIC(Alarm_Pure_Steam_High_Temperature_Ack) ,XIC(S:FS) ]OTU(Alarm_Pure_Steam_High_Temperature);
   28: XIC(AI_R_2_0_Pure_Steam_Temperature.Fault)TON(Alarm_Pure_Steam_Temp_Error_Timer,?,?);
